// Verrouillages d'une station (docs/04 § 4) : 0 si autorisé, sinon n° du verrouillage violé
INTERFACE I_InterlockProvider

METHOD Check : INT
VAR_INPUT
    nLocalId : UINT;
    nAction : UINT;
END_VAR
END_METHOD

END_INTERFACE

(* stored: Version 1.1.0.1, ProductVersion 3.1.4024.12
   Itf I_InterlockProvider: Id {7114bd0c-a703-5ab6-b124-d008ab6b5348}
   Method Check: Id {8714eae5-9a4c-5d0e-a74a-4d781a25dc30} *)
